(*
SPDX-FileCopyrightText: © 2026 Oleksandr Tiutyk <trofimich@gmail.com>
SPDX-License-Identifier: MIT
License: https://opensource.org/license/mit
*)

(*!
<summary>Serializes live PLC structures to JSON and restores them from JSON.</summary>
<description>
Supports live PLC structures with native type information; dynamically created structures are not supported.
ByVarInfo methods require an explicit PVOID address; descriptor ByteAddress is ignored to preserve pointer width.
Application method calls and property access belong to one owner task per instance. Instances are not
thread-safe and do not support reentry: a callback must not call methods or access properties of the
serializer whose operation is still active, directly or indirectly. Use a separate instance and separate
buffers for another task or nested conversion. Ownership is a caller precondition, not a runtime check or
lock; Try does not make an ownership violation safe or guarantee its detection as FALSE. Keep source data
stable and destination storage exclusive for the entire call, including callbacks. Separate serializer
instances do not synchronize shared application data. Stateful extenders require their own ownership
discipline; sharing an extender must not introduce concurrent state access. Borrows input, output and optional
callbacks for each call. Throwing methods report invalid arguments and native failures through framework
exceptions. Try methods return FALSE directly for rejected arguments or reported native failures and contain
exceptions from native calls or callbacks; partial effects are not rolled back. Try methods use the shared
native conversion helpers, not overrides of the throwing methods or their protected helpers. JSON text uses
native UTF-8 encoding; capacity and copy sizes count bytes. Instances must not be copied by value. The caller
provides cyclic-task exception cleanup and RaiseIfAllocationFailed at the task boundary, outside Try and
recoverable handlers. Try methods do not clear terminal allocation state. Ownership examples and future
shared-service guidance: Guides/JsonAndEventLoggerOwnership.md in the repository.
</description>
*)

{attribute 'no_explicit_call' := 'Direct call is not allowed'}
FUNCTION_BLOCK AutomaticJsonSerializer EXTENDS TOF_Core.Object
VAR_STAT
	//! <summary>Class name shared by all instances of this function block.</summary>
	{attribute 'hide'} 
	_ClassName : STRING := __POUNAME();
END_VAR
VAR
	_JsonSaxWriter : Tc3_JsonXml.FB_JsonSaxWriter;
	_JsonDataTypeWriter : Tc3_JsonXml.FB_JsonReadWriteDatatype;
END_VAR

(*!
<summary>Provides the concrete serializer class name.</summary>
<description>Borrows read-only instance storage that remains valid for the instance lifetime.</description>
*)
{attribute 'monitoring' := 'call'}
PROPERTY ClassName : REFERENCE TO STRING
GET
ClassName REF= _ClassName;
END_GET
END_PROPERTY

(*!
<summary>Serializes a PLC structure into caller-owned JSON storage.</summary>
<description>
Uses native symbol lookup for the source type; dynamically created structures are not supported. Single-field
structures have native lookup limitations; use ByVarInfo to supply the type explicitly. Borrows
source, destination and optional extender for the call. The destination must be writable and have at least
JSON_DOCUMENT capacity. Invalid source arguments and reported native failures raise framework exceptions;
extender exceptions propagate. Output and callback effects are not rolled back on failure. Exception transport
and cleanup require the caller's cyclic-task boundary. CopyDocument returning zero or a nonzero HRESULT raises
an exception; jsonSize is not usable on failure.
</description>
<param name="sourceStructure">Live PLC structure with type information available to native symbol lookup.</param>
<param name="extender">
Optional callback invoked before and after writing the structure value; zero skips both calls.
</param>
<param name="targetJson">Writable output storage with at least 25000 bytes of text capacity plus the terminator.</param>
<param name="jsonSize">
Byte count reported by CopyDocument, including the terminator on a successful copy; use only after normal
completion.
</param>
*)
METHOD Serialize
VAR_INPUT
	sourceStructure : ANY;
	extender : IJsonExtender := 0;
END_VAR
VAR_IN_OUT
	targetJson : TOF_Core.JSON_DOCUMENT;
END_VAR
VAR_OUTPUT
	jsonSize : UDINT; 
END_VAR
InternalSerialize(
	sourceStructure := sourceStructure,
	extender := extender,
	targetJson := targetJson,
	jsonSize => jsonSize
);
END_METHOD

(*!
<summary>Serializes a PLC structure described by VAR_INFO into caller-owned JSON storage.</summary>
<description>
The descriptor type and byte-aligned size must match sourceStructureAddress. ByteAddress is ignored.
Dynamically created structures are not supported. Borrows source, destination and optional extender for the call. The
destination must be writable and have at least JSON_DOCUMENT capacity. Invalid source arguments and reported
native failures raise framework exceptions; extender exceptions propagate. Output and callback effects are not
rolled back on failure. Exception transport and cleanup require the caller's cyclic-task boundary.
CopyDocument returning zero or a nonzero HRESULT raises an exception; jsonSize is not usable on failure.
</description>
<param name="sourceStructureAddress">
Required address from ADR of the live source structure, borrowed for this call. Must match the descriptor.
Zero is rejected; no address is recovered from ByteAddress or ByteOffset.
</param>
<param name="sourceStructureVarInfo">
Descriptor whose TypeName and BitSize describe the source structure; ByteAddress is ignored.
</param>
<param name="extender">
Optional callback invoked before and after writing the structure value; zero skips both calls.
</param>
<param name="targetJson">Writable output storage with at least 25000 bytes of text capacity plus the terminator.</param>
<param name="jsonSize">
Byte count reported by CopyDocument, including the terminator on a successful copy; use only after normal
completion.
</param>
*)
METHOD SerializeByVarInfo
VAR_INPUT
	sourceStructureVarInfo : __SYSTEM.VAR_INFO;
	sourceStructureAddress : PVOID;
	extender : IJsonExtender := 0;
END_VAR
VAR_IN_OUT
	targetJson : TOF_Core.JSON_DOCUMENT;
END_VAR
VAR_OUTPUT
	jsonSize : UDINT; 
END_VAR
VAR
	formattedExceptionMessage : TOF_Core.ERROR_MESSAGE;

	
	errorCode : HRESULT;
END_VAR
IF sourceStructureAddress = TOF_Core.Memory.NULL_ADDRESS THEN
	TOF_Core.Exceptions.ThrowArgumentNotSpecified(
		sourceNamespaceName := NamespaceName,
		sourceClassName := ClassName,
		sourcePOUName := __POUNAME(),
		sourcePosition := __POSITION(),
		argumentName := 'sourceStructureAddress'
	);
END_IF

IF sourceStructureVarInfo.TypeClass <> __SYSTEM.TYPE_CLASS.TYPE_USERDEF THEN
	TOF_Core.Exceptions.ThrowArgumentTypeClassNotSupported(
		sourceNamespaceName := NamespaceName,
		sourceClassName := ClassName,
		sourcePOUName := __POUNAME(),
		sourcePosition := __POSITION(),
		argumentName := 'sourceStructureVarInfo',
		argumentType := sourceStructureVarInfo.TypeClass
	);
END_IF

// VAR_INFO sizes are in bits; the caller supplies a byte-aligned structure descriptor.
IF NOT writeStructureJson(
	structureTypeName := sourceStructureVarInfo.TypeName,
	structureAddress := sourceStructureAddress,
	structureSize := TO_UDINT(sourceStructureVarInfo.BitSize / 8),
	extender := extender,
	targetJson := targetJson,
	jsonSize => jsonSize,
	errorCode => errorCode,
	errorMessage => formattedExceptionMessage
)
THEN
	TOF_Core.Exceptions.ThrowStandard(
		sourceNamespaceName := NamespaceName,
		sourceClassName := ClassName,
		sourcePOUName := __POUNAME(),
		sourcePosition := __POSITION(),
		message := formattedExceptionMessage,
		errorCode := TO_UDINT(errorCode)
	);
END_IF
END_METHOD

{attribute 'monitoring' := 'call'}
(*!
<summary>Gets or sets the native writer's maximum number of fractional decimal places.</summary>
<description>
The native writer determines which DINT values it supports; this property does not clamp the value. The setter
requires a zero HRESULT from SetMaxDecimalPlaces. A nonzero HRESULT raises a framework exception because
assignment has no failure result. The native error code is retained in the exception. No rollback of the
native setting is guaranteed on failure; the getter reads the writer's current setting. The caller handles the
exception and provides cyclic-task exception cleanup and the terminal allocation-failure boundary.
</description>
*)
PROPERTY DecimalPlaces : DINT
GET
DecimalPlaces := _JsonSaxWriter.GetMaxDecimalPlaces();
END_GET
SET
VAR
	errorCode : HRESULT;
END_VAR
errorCode := _JsonSaxWriter.SetMaxDecimalPlaces(decimalPlaces := DecimalPlaces);

IF errorCode <> TOF_Core.SignedInt32.ZERO THEN
	TOF_Core.Exceptions.ThrowStandard(
		sourceNamespaceName := NamespaceName,
		sourceClassName := ClassName,
		sourcePOUName := __POUNAME(),
		sourcePosition := __POSITION(),
		message := "Can't set JSON writer decimal places",
		errorCode := TO_UDINT(errorCode)
	);
END_IF
END_SET
END_PROPERTY

(*!
<summary>Populates a PLC structure from JSON using the type supplied by VAR_INFO.</summary>
<description>
TypeName and byte-aligned BitSize must describe the live, writable structure at targetStructureAddress.
ByteAddress is ignored. Uses the supplied TypeName directly, avoiding ambiguous address-based type lookup
for single-field structures. The type
must be available to the native JSON converter; support for dynamically created structures is not implied.
Borrows the JSON and destination for this call. A zero address, an unsupported type class or a reported native
conversion failure raises a framework exception. Conversion requires both a TRUE SetSymbolFromJson result and
a zero HRESULT. Destination fields may already have changed on failure; writes are not rolled back. The caller
provides cyclic-task exception cleanup and the terminal allocation-failure boundary.
</description>
<param name="json">JSON text to read without modification.</param>
<param name="targetStructureAddress">
Required address from ADR of the live target structure, borrowed for this call. Must match the descriptor.
Zero is rejected; no address is recovered from ByteAddress or ByteOffset.
</param>
<param name="targetStructureVarInfo">
Consistent descriptor of the destination structure, including its explicit TypeName.
</param>
*)
METHOD DeserializeByVarInfo
VAR_IN_OUT CONSTANT
	json : TOF_Core.JSON_DOCUMENT;	
END_VAR
VAR_INPUT
	targetStructureVarInfo : __SYSTEM.VAR_INFO;
	targetStructureAddress : PVOID;
END_VAR
VAR
	
	errorCode : HRESULT;
END_VAR
IF targetStructureAddress = TOF_Core.Memory.NULL_ADDRESS THEN
	TOF_Core.Exceptions.ThrowArgumentNotSpecified(
		sourceNamespaceName := NamespaceName,
		sourceClassName := ClassName,
		sourcePOUName := __POUNAME(),
		sourcePosition := __POSITION(),
		argumentName := 'targetStructureAddress'
	);
END_IF

IF targetStructureVarInfo.TypeClass <> __SYSTEM.TYPE_CLASS.TYPE_USERDEF THEN
	TOF_Core.Exceptions.ThrowArgumentTypeClassNotSupported(
		sourceNamespaceName := NamespaceName,
		sourceClassName := ClassName,
		sourcePOUName := __POUNAME(),
		sourcePosition := __POSITION(),
		argumentName := 'targetStructureVarInfo',
		argumentType := targetStructureVarInfo.TypeClass
	);
END_IF

// VAR_INFO sizes are in bits; the caller supplies a byte-aligned structure descriptor.
IF NOT readStructureJson(
	json := json,
	structureTypeName := targetStructureVarInfo.TypeName,
	structureAddress := targetStructureAddress,
	structureSize := TO_UDINT(targetStructureVarInfo.BitSize / 8),
	errorCode => errorCode
)
THEN
	TOF_Core.Exceptions.ThrowStandard(
		sourceNamespaceName := NamespaceName,
		sourceClassName := ClassName,
		sourcePOUName := __POUNAME(),
		sourcePosition := __POSITION(),
		message := "Can't fill target structure by specified json document",
		errorCode := TO_UDINT(errorCode)
	);
END_IF
END_METHOD

(*!
<summary>Populates a PLC structure from JSON using native address-based type lookup.</summary>
<description>
Borrows the JSON and a live, writable structure for the call; dynamically created structures are not
supported. Native type lookup has limitations for single-field structures. Invalid arguments, reported lookup
failures, a FALSE SetSymbolFromJson result or a nonzero conversion HRESULT raise framework exceptions.
Destination fields may already have changed on failure; writes are not rolled back. The caller provides
cyclic-task exception cleanup and the terminal allocation-failure boundary.
</description>
<param name="json">JSON text to read without modification.</param>
<param name="targetStructure">
Live destination structure with type information available to native symbol lookup.
</param>
*)
METHOD Deserialize
VAR_IN_OUT CONSTANT
	json : TOF_Core.JSON_DOCUMENT;	
END_VAR
VAR_INPUT
	targetStructure : ANY;
END_VAR
InternalDeserialize(json := json, targetStructure := targetStructure);
END_METHOD

(*!
<summary>Serializes a structure using its ANY descriptor and native symbol lookup.</summary>
<description>
The descriptor must identify a live structure with matching address and size; dynamically created structures
are not supported. Native address lookup has limitations for single-field structures. Borrows source,
destination and optional extender for the call. The destination must be writable and have at least
JSON_DOCUMENT capacity. Invalid source arguments and reported native failures raise framework exceptions;
extender exceptions propagate. Output and callback effects are not rolled back on failure. Overrides must
preserve destination capacity and borrowing requirements. This protected hook serves the throwing ANY API;
TrySerialize does not dispatch through it. Exception transport and cleanup require the caller's
cyclic-task boundary. CopyDocument returning zero or a nonzero HRESULT raises an exception; jsonSize is not
usable on failure.
</description>
<param name="sourceStructure">ANY descriptor for the source structure.</param>
<param name="extender">
Optional callback invoked before and after writing the structure value; zero skips both calls.
</param>
<param name="targetJson">Writable output storage with at least 25000 bytes of text capacity plus the terminator.</param>
<param name="jsonSize">
Byte count reported by CopyDocument, including the terminator on a successful copy; use only after normal
completion.
</param>
*)
METHOD PROTECTED InternalSerialize
VAR_INPUT
	sourceStructure : __SYSTEM.AnyType;
	extender : IJsonExtender := 0;
END_VAR
VAR_IN_OUT
	targetJson : TOF_Core.JSON_DOCUMENT;
END_VAR
VAR_OUTPUT
	jsonSize : UDINT; 
END_VAR
VAR
	formattedExceptionMessage : TOF_Core.ERROR_MESSAGE;

	
	structureTypeName : STRING;	 
	errorCode : HRESULT;
END_VAR
IF sourceStructure.pValue = TOF_Core.Memory.NULL_ADDRESS THEN
	TOF_Core.Exceptions.ThrowArgumentNotSpecified(
		sourceNamespaceName := NamespaceName,
		sourceClassName := ClassName,
		sourcePOUName := __POUNAME(),
		sourcePosition := __POSITION(),
		argumentName := 'sourceStructure'
	);
END_IF

IF sourceStructure.TypeClass <> __SYSTEM.TYPE_CLASS.TYPE_USERDEF THEN
	TOF_Core.Exceptions.ThrowArgumentTypeClassNotSupported(
		sourceNamespaceName := NamespaceName,
		sourceClassName := ClassName,
		sourcePOUName := __POUNAME(),
		sourcePosition := __POSITION(),
		argumentName := 'sourceStructure',
		argumentType := sourceStructure.TypeClass
	);
END_IF

structureTypeName := _JsonDataTypeWriter.GetDatatypeNameByAddress(
	nData := TO_UDINT(sourceStructure.diSize),
	pData := sourceStructure.pValue,
	hrErrorCode => errorCode
);

IF errorCode <> TOF_Core.SignedInt32.ZERO THEN
	TOF_Core.Exceptions.ThrowStandard(
		sourceNamespaceName := NamespaceName,
		sourceClassName := ClassName,
		sourcePOUName := __POUNAME(),
		sourcePosition := __POSITION(),
		message := "Can't get structure type of the source structure",
		errorCode := TO_UDINT(errorCode)
	);
END_IF

IF NOT writeStructureJson(
	structureTypeName := structureTypeName,
	structureAddress := sourceStructure.pValue,
	structureSize := TO_UDINT(sourceStructure.diSize),
	extender := extender,
	targetJson := targetJson,
	jsonSize => jsonSize,
	errorCode => errorCode,
	errorMessage => formattedExceptionMessage
)
THEN
	TOF_Core.Exceptions.ThrowStandard(
		sourceNamespaceName := NamespaceName,
		sourceClassName := ClassName,
		sourcePOUName := __POUNAME(),
		sourcePosition := __POSITION(),
		message := formattedExceptionMessage,
		errorCode := TO_UDINT(errorCode)
	);
END_IF
END_METHOD

(*!
<summary>Deserializes JSON into the structure identified by an ANY descriptor.</summary>
<description>
The descriptor must identify a live, writable structure with matching address and size; dynamically created
structures are not supported. Native address-based type lookup has limitations for single-field structures.
Borrows the JSON and destination for the call. Invalid arguments, reported lookup failures, a FALSE
SetSymbolFromJson result or a nonzero conversion HRESULT raise framework exceptions. Partial destination
writes are not rolled back. Overrides must preserve borrowing and failure reporting requirements. This
protected hook serves the throwing ANY API; TryDeserialize does not dispatch through it. The caller
provides cyclic-task exception cleanup and the terminal allocation-failure boundary.
</description>
<param name="json">JSON text to read without modification.</param>
<param name="targetStructure">ANY descriptor for the live destination structure.</param>
*)
METHOD PROTECTED InternalDeserialize
VAR_IN_OUT CONSTANT
	json : TOF_Core.JSON_DOCUMENT;	
END_VAR
VAR_INPUT
	targetStructure : __SYSTEM.AnyType;
END_VAR
VAR
	
	structureTypeName : STRING;	 
	errorCode : HRESULT;
END_VAR
IF targetStructure.pValue = TOF_Core.Memory.NULL_ADDRESS THEN
	TOF_Core.Exceptions.ThrowArgumentNotSpecified(
		sourceNamespaceName := NamespaceName,
		sourceClassName := ClassName,
		sourcePOUName := __POUNAME(),
		sourcePosition := __POSITION(),
		argumentName := 'targetStructure'
	);
END_IF

IF targetStructure.TypeClass <> __SYSTEM.TYPE_CLASS.TYPE_USERDEF THEN
	TOF_Core.Exceptions.ThrowArgumentTypeClassNotSupported(
		sourceNamespaceName := NamespaceName,
		sourceClassName := ClassName,
		sourcePOUName := __POUNAME(),
		sourcePosition := __POSITION(),
		argumentName := 'targetStructure',
		argumentType := targetStructure.TypeClass
	);
END_IF

structureTypeName := _JsonDataTypeWriter.GetDatatypeNameByAddress(
	nData := TO_UDINT(targetStructure.diSize),
	pData := targetStructure.pValue,
	hrErrorCode => errorCode
);

IF errorCode <> TOF_Core.SignedInt32.ZERO THEN
	TOF_Core.Exceptions.ThrowStandard(
		sourceNamespaceName := NamespaceName,
		sourceClassName := ClassName,
		sourcePOUName := __POUNAME(),
		sourcePosition := __POSITION(),
		message := "Can't get structure type of the target structure",
		errorCode := TO_UDINT(errorCode)
	);
END_IF

IF NOT readStructureJson(
	json := json,
	structureTypeName := structureTypeName,
	structureAddress := targetStructure.pValue,
	structureSize := TO_UDINT(targetStructure.diSize),
	errorCode => errorCode
)
THEN
	TOF_Core.Exceptions.ThrowStandard(
		sourceNamespaceName := NamespaceName,
		sourceClassName := ClassName,
		sourcePOUName := __POUNAME(),
		sourcePosition := __POSITION(),
		message := "Can't fill target structure by specified json document",
		errorCode := TO_UDINT(errorCode)
	);
END_IF
END_METHOD

(*!
<summary>Provides the compiler-initialized library namespace.</summary>
<description>Borrows read-only library storage; no allocation or ownership transfer occurs.</description>
*)
{attribute 'monitoring' := 'call'}
PROPERTY NamespaceName : REFERENCE TO STRING
GET
NamespaceName REF= CurrentNamespace.Name;
END_GET
END_PROPERTY

(*!
<summary>Reads JSON into a validated structure and reports the native conversion result.</summary>
<description>
Callers validate the descriptor before entry. Borrows the JSON, type name and destination for this call.
Returns FALSE for a native FALSE result or nonzero HRESULT without creating exceptions. Native exceptions
propagate to the throwing caller or the public Try boundary. Checks fatal allocation state before conversion
and before reporting success, raising a contained terminal failure without constructing an exception object.
The Try boundary converts that failure to FALSE. Partial destination writes are not rolled back.
</description>
<param name="json">JSON text to read without modification.</param>
<param name="structureTypeName">Native type name matching the destination structure.</param>
<param name="structureAddress">Address of the validated writable destination.</param>
<param name="structureSize">Destination structure size in bytes.</param>
<param name="errorCode">Native conversion HRESULT, interpreted together with the BOOL result.</param>
*)
METHOD PRIVATE readStructureJson : BOOL
VAR_IN_OUT CONSTANT
	json : TOF_Core.JSON_DOCUMENT;
	structureTypeName : STRING;
END_VAR
VAR_INPUT
	structureAddress : PVOID;
	structureSize : UDINT;
END_VAR
VAR_OUTPUT
	errorCode : HRESULT;
END_VAR
TOF_Core.DynamicMemoryManager.RaiseIfAllocationFailed();

IF NOT _JsonDataTypeWriter.SetSymbolFromJson(
		sJson := json,
		sDatatype := structureTypeName,
		nData := structureSize,
		pData := structureAddress,
		hrErrorCode => errorCode
	)
	OR_ELSE errorCode <> TOF_Core.SignedInt32.ZERO
THEN
	RETURN;
END_IF

TOF_Core.DynamicMemoryManager.RaiseIfAllocationFailed();
readStructureJson := TRUE;
END_METHOD

(*!
<summary>Reports the complete instance size in bytes.</summary>
<description>Uses XSIZEOF; separately allocated native resources are not included.</description>
*)
{attribute 'monitoring' := 'call'}
PROPERTY SelfSize : ULINT
GET
SelfSize := XSIZEOF(THIS^);
END_GET
END_PROPERTY

{attribute 'TcRpcEnable':='1'}
(*!
<summary>Attempts to serialize a PLC structure to JSON.</summary>
<description>
Returns FALSE directly for a null address, an unsupported type class or a reported native failure, including a
zero CopyDocument result, without creating a framework exception. Contains native and callback exceptions.
Uses the shared conversion helper rather than the protected throwing hook. Use JSON and jsonSize only on TRUE;
partial writes and callback effects are not rolled back. Each subsequent conversion attempts to reset the
writer before callbacks. Borrows live source and writable destination storage. Does not clear terminal allocation state; the
caller provides exception cleanup and RaiseIfAllocationFailed at the task boundary outside Try and recoverable
handlers. Returns FALSE when fatal allocation state is observed on entry or after nested calls; a contained
allocation failure is not a successful conversion. The application-wide latch remains set.
</description>
<param name="sourceStructure">
Live PLC structure supported by native symbol lookup; dynamically created structures are not supported.
Single-field structures have native lookup limitations; use ByVarInfo to supply the type explicitly.
</param>
<param name="extender">
Optional callback invoked before and after writing the structure value; borrowed for the call.
</param>
<param name="targetJson">
Writable output storage with at least 25000 bytes of text capacity plus the terminator; borrowed for the call.
</param>
<param name="jsonSize">
Byte count reported by CopyDocument, including the terminator on a successful copy; use only on TRUE.
</param>
*)
METHOD TrySerialize : BOOL
VAR_INPUT
	sourceStructure : ANY;
	extender : IJsonExtender := 0;
END_VAR
VAR_IN_OUT
	targetJson : TOF_Core.JSON_DOCUMENT;
END_VAR
VAR_OUTPUT
	jsonSize : UDINT; 
END_VAR
VAR
	structureTypeName : STRING;
	errorCode : HRESULT;
END_VAR
__TRY

	IF TOF_Core.DynamicMemoryManager.HasAllocationFailed THEN
		RETURN;
	END_IF

	IF sourceStructure.pValue = TOF_Core.Memory.NULL_ADDRESS
		OR_ELSE sourceStructure.TypeClass <> __SYSTEM.TYPE_CLASS.TYPE_USERDEF
	THEN
		RETURN;
	END_IF

	structureTypeName := _JsonDataTypeWriter.GetDatatypeNameByAddress(
		nData := TO_UDINT(sourceStructure.diSize),
		pData := sourceStructure.pValue,
		hrErrorCode => errorCode
	);

	IF errorCode <> TOF_Core.SignedInt32.ZERO THEN
		RETURN;
	END_IF

	TrySerialize := writeStructureJson(
		structureTypeName := structureTypeName,
		structureAddress := sourceStructure.pValue,
		structureSize := TO_UDINT(sourceStructure.diSize),
		extender := extender,
		targetJson := targetJson,
		jsonSize => jsonSize
	);

	IF TOF_Core.DynamicMemoryManager.HasAllocationFailed THEN
		TrySerialize := FALSE;
	END_IF

__CATCH
	TrySerialize := FALSE;
__ENDTRY
END_METHOD

(*!
<summary>Attempts to serialize a PLC structure to JSON.</summary>
<description>
Returns FALSE directly for a null address, an unsupported type class or a reported native failure, including a
zero CopyDocument result, without creating a framework exception. Contains native and callback exceptions.
Uses the shared conversion helper rather than the throwing ByVarInfo method. Use JSON and jsonSize only on
TRUE; partial writes and callback effects are not rolled back. Each subsequent conversion attempts to reset
the writer before callbacks. Borrows live source and writable destination storage. Does not clear terminal allocation
state; the caller provides exception cleanup and RaiseIfAllocationFailed at the task boundary outside Try and
recoverable handlers. Returns FALSE when fatal allocation state is observed on entry or after nested calls; a contained
allocation failure is not a successful conversion. The application-wide latch remains set.
</description>
<param name="sourceStructureAddress">
Required address from ADR of the live source structure, borrowed for this call. Must match the descriptor.
Zero is rejected; no address is recovered from ByteAddress or ByteOffset.
</param>
<param name="sourceStructureVarInfo">
Descriptor with matching TypeName and byte-aligned BitSize for sourceStructureAddress; ByteAddress is ignored.
Dynamically created structures are not supported.
</param>
<param name="extender">
Optional callback invoked before and after writing the structure value; borrowed for the call.
</param>
<param name="targetJson">
Writable output storage with at least 25000 bytes of text capacity plus the terminator; borrowed for the call.
</param>
<param name="jsonSize">
Byte count reported by CopyDocument, including the terminator on a successful copy; use only on TRUE.
</param>
*)
METHOD TrySerializeByVarInfo : BOOL
VAR_INPUT
	sourceStructureVarInfo : __SYSTEM.VAR_INFO;
	sourceStructureAddress : PVOID;
	extender : IJsonExtender := 0;
END_VAR
VAR_IN_OUT
	targetJson : TOF_Core.JSON_DOCUMENT;
END_VAR
VAR_OUTPUT
	jsonSize : UDINT; 
END_VAR
__TRY

	IF TOF_Core.DynamicMemoryManager.HasAllocationFailed THEN
		RETURN;
	END_IF

	IF sourceStructureAddress = TOF_Core.Memory.NULL_ADDRESS
		OR_ELSE sourceStructureVarInfo.TypeClass <> __SYSTEM.TYPE_CLASS.TYPE_USERDEF
	THEN
		RETURN;
	END_IF

	// VAR_INFO sizes are in bits; the descriptor must be byte-aligned.
	TrySerializeByVarInfo := writeStructureJson(
		structureTypeName := sourceStructureVarInfo.TypeName,
		structureAddress := sourceStructureAddress,
		structureSize := TO_UDINT(sourceStructureVarInfo.BitSize / 8),
		extender := extender,
		targetJson := targetJson,
		jsonSize => jsonSize
	);

	IF TOF_Core.DynamicMemoryManager.HasAllocationFailed THEN
		TrySerializeByVarInfo := FALSE;
	END_IF

__CATCH
	TrySerializeByVarInfo := FALSE;
__ENDTRY
END_METHOD

(*!
<summary>Attempts to populate a PLC structure from JSON using the type supplied by VAR_INFO.</summary>
<description>
Uses the supplied TypeName directly without address-based type lookup. TypeName and byte-aligned BitSize must
describe the live, writable structure at targetStructureAddress, with its type available to the native converter.
ByteAddress is ignored.
Returns FALSE directly for a null address, an unsupported type class, a FALSE native conversion result or a
nonzero HRESULT, without creating a framework exception. Contains native exceptions. Uses the shared
conversion helper rather than the throwing ByVarInfo method. Partial destination writes are not rolled back.
Borrows the JSON and destination for this call. Does not clear terminal allocation state; the caller provides
exception cleanup and RaiseIfAllocationFailed at the task boundary outside Try and recoverable handlers.
Returns FALSE when fatal allocation state is observed on entry or after nested calls; a contained
allocation failure is not a successful conversion. The application-wide latch remains set.
</description>
<param name="json">JSON text to read without modification.</param>
<param name="targetStructureAddress">
Required address from ADR of the live target structure, borrowed for this call. Must match the descriptor.
Zero is rejected; no address is recovered from ByteAddress or ByteOffset.
</param>
<param name="targetStructureVarInfo">
Consistent descriptor of the destination structure, including its explicit TypeName.
</param>
*)
METHOD TryDeserializeByVarInfo : BOOL
VAR_IN_OUT CONSTANT
	json : TOF_Core.JSON_DOCUMENT;	
END_VAR
VAR_INPUT
	targetStructureVarInfo : __SYSTEM.VAR_INFO;
	targetStructureAddress : PVOID;
END_VAR
__TRY

	IF TOF_Core.DynamicMemoryManager.HasAllocationFailed THEN
		RETURN;
	END_IF

	IF targetStructureAddress = TOF_Core.Memory.NULL_ADDRESS
		OR_ELSE targetStructureVarInfo.TypeClass <> __SYSTEM.TYPE_CLASS.TYPE_USERDEF
	THEN
		RETURN;
	END_IF

	// VAR_INFO sizes are in bits; the descriptor must be byte-aligned.
	TryDeserializeByVarInfo := readStructureJson(
		json := json,
		structureTypeName := targetStructureVarInfo.TypeName,
		structureAddress := targetStructureAddress,
		structureSize := TO_UDINT(targetStructureVarInfo.BitSize / 8)
	);

	IF TOF_Core.DynamicMemoryManager.HasAllocationFailed THEN
		TryDeserializeByVarInfo := FALSE;
	END_IF

__CATCH
	TryDeserializeByVarInfo := FALSE;
__ENDTRY
END_METHOD

(*!
<summary>Attempts to populate a PLC structure from JSON.</summary>
<description>
Uses native address-based type lookup, with its limitations for single-field structures; dynamically created
structures are not supported. Returns FALSE directly for a null address, an unsupported type class, a reported
lookup failure, a FALSE native conversion result or a nonzero conversion HRESULT, without creating a framework
exception. Contains native exceptions. Uses the shared conversion helper rather than the protected throwing
hook. Partial destination writes are not rolled back. Borrows JSON and live, writable destination storage for
this call. Does not clear terminal allocation state; the caller provides exception cleanup and
RaiseIfAllocationFailed at the task boundary outside Try and recoverable handlers.
Returns FALSE when fatal allocation state is observed on entry or after nested calls; a contained
allocation failure is not a successful conversion. The application-wide latch remains set.
</description>
<param name="json">JSON text to read without modification.</param>
<param name="targetStructure">
Live destination structure with type information available to native symbol lookup.
</param>
*)
METHOD TryDeserialize : BOOL
VAR_IN_OUT CONSTANT
	json : TOF_Core.JSON_DOCUMENT;	
END_VAR
VAR_INPUT
	targetStructure : ANY;
END_VAR
VAR
	structureTypeName : STRING;
	errorCode : HRESULT;
END_VAR
__TRY

	IF TOF_Core.DynamicMemoryManager.HasAllocationFailed THEN
		RETURN;
	END_IF

	IF targetStructure.pValue = TOF_Core.Memory.NULL_ADDRESS
		OR_ELSE targetStructure.TypeClass <> __SYSTEM.TYPE_CLASS.TYPE_USERDEF
	THEN
		RETURN;
	END_IF

	structureTypeName := _JsonDataTypeWriter.GetDatatypeNameByAddress(
		nData := TO_UDINT(targetStructure.diSize),
		pData := targetStructure.pValue,
		hrErrorCode => errorCode
	);

	IF errorCode <> TOF_Core.SignedInt32.ZERO THEN
		RETURN;
	END_IF

	TryDeserialize := readStructureJson(
		json := json,
		structureTypeName := structureTypeName,
		structureAddress := targetStructure.pValue,
		structureSize := TO_UDINT(targetStructure.diSize)
	);

	IF TOF_Core.DynamicMemoryManager.HasAllocationFailed THEN
		TryDeserialize := FALSE;
	END_IF

__CATCH
	TryDeserialize := FALSE;
__ENDTRY
END_METHOD

(*!
<summary>Writes a validated structure and optional extensions to caller-owned JSON storage.</summary>
<description>
Callers validate the structure descriptor before entry. Borrows all arguments for this call and resets the
writer before invoking callbacks. A nonzero ResetDocument HRESULT returns FALSE before any hook or copy.
Returns FALSE for reported native failures without creating exceptions; native or callback exceptions propagate
to the throwing caller or the public Try boundary. Checks fatal allocation state before native work, after
successful native steps and after each hook. A contained terminal failure is raised again without allocating
an exception object; the Try boundary converts it to FALSE. No output, writer or callback effects are rolled
back. Each later write attempts to reset the writer again. On FALSE, errorMessage describes the failed native
step and errorCode retains its HRESULT without substitution.
</description>
<param name="structureTypeName">Native type name matching the live source structure.</param>
<param name="structureAddress">Address of the validated source structure.</param>
<param name="structureSize">Source structure size in bytes.</param>
<param name="extender">Optional callbacks around the structure value.</param>
<param name="targetJson">Writable storage with JSON_DOCUMENT capacity, including its terminator.</param>
<param name="jsonSize">Copied byte count including the terminator; meaningful only on TRUE.</param>
<param name="errorCode">Native HRESULT of the failed step on FALSE.</param>
<param name="errorMessage">Diagnostic for the failed step on FALSE.</param>
*)
METHOD PRIVATE writeStructureJson : BOOL
VAR_IN_OUT CONSTANT
	structureTypeName : STRING;
END_VAR
VAR_INPUT
	structureAddress : PVOID;
	structureSize : UDINT;
	extender : IJsonExtender;
END_VAR
VAR_IN_OUT
	targetJson : TOF_Core.JSON_DOCUMENT;
END_VAR
VAR_OUTPUT
	jsonSize : UDINT;
	errorCode : HRESULT;
	errorMessage : WSTRING(255);
END_VAR
TOF_Core.DynamicMemoryManager.RaiseIfAllocationFailed();
errorCode := _JsonSaxWriter.ResetDocument();
TOF_Core.DynamicMemoryManager.RaiseIfAllocationFailed();

IF errorCode <> TOF_Core.SignedInt32.ZERO THEN
	errorMessage := "Can't reset JSON writer before structure serialization";
	RETURN;
END_IF

IF extender <> 0 THEN
	extender.WritePrefix(jsonSaxWriter := _JsonSaxWriter);
	TOF_Core.DynamicMemoryManager.RaiseIfAllocationFailed();
END_IF

IF NOT _JsonDataTypeWriter.AddJsonValueFromSymbol(
		fbWriter := _JsonSaxWriter,
		sDatatype := structureTypeName,
		nData := structureSize,
		pData := structureAddress,
		hrErrorCode => errorCode
	)
	OR_ELSE errorCode <> TOF_Core.SignedInt32.ZERO
THEN
	errorMessage := TOF_Core.WideStrings.Concat255(
		"Can't generate JSON representation from the symbol of type '",
		TO_WSTRING(structureTypeName),
		"'"
	);
	RETURN;
END_IF

TOF_Core.DynamicMemoryManager.RaiseIfAllocationFailed();

IF extender <> 0 THEN
	extender.WriteSuffix(jsonSaxWriter := _JsonSaxWriter);
	TOF_Core.DynamicMemoryManager.RaiseIfAllocationFailed();
END_IF

jsonSize := _JsonSaxWriter.CopyDocument(
	pDoc := targetJson,
	nDoc := SIZEOF(targetJson),
	hrErrorCode => errorCode
);

IF jsonSize = TOF_Core.UnsignedInt32.MIN_VALUE OR_ELSE errorCode <> TOF_Core.SignedInt32.ZERO THEN
	errorMessage := TOF_Core.WideStrings.Concat255(
		"Can't fill JSON from the symbol of type '",
		TO_WSTRING(structureTypeName),
		"'"
	);
	RETURN;
END_IF

TOF_Core.DynamicMemoryManager.RaiseIfAllocationFailed();
writeStructureJson := TRUE;
END_METHOD

END_FUNCTION_BLOCK

(* stored: Version 1.1.0.1
   POU AutomaticJsonSerializer: Id {a4623321-e5e2-4514-b5b7-6f50c93efdb9}, SpecialFunc None
   Folder Service memebers: Id {ac3ba484-d0b1-4d7e-b557-cd243c8b8997}
   Property ClassName: Id {0ef034e0-c59c-400d-8910-5199a1e43c28}
   Get Get: Id {7d8e441f-d9e1-4fe6-a84f-2d3a88ae1b83}
   Method Serialize: Id {defd30bb-3636-4b3d-a29d-4ee5f3966212}
   Method SerializeByVarInfo: Id {d6f652b9-17a4-4ec4-936c-676a73e01a2d}
   Property DecimalPlaces: Id {856a998f-c63b-4bfb-be2d-ebc0ce7cf745}
   Get Get: Id {94eff383-c1b9-45b7-8cbb-da0c6c3a2aac}
   Set Set: Id {e5e3c1bb-4425-43f2-a416-2b4fee3a3ddc}
   Method DeserializeByVarInfo: Id {3b0559f7-3cc9-4407-b03c-9992acf72583}
   Method Deserialize: Id {b53042c3-1eea-4151-a973-f56939241dea}
   Method InternalSerialize: Id {828ddc06-4e4b-4f22-bd8f-3234f73fd728}
   Method InternalDeserialize: Id {cd668581-fbff-4bb3-b0d3-914c47132fdf}
   Property NamespaceName: Id {7371ecef-1936-4268-af0d-813ed5877183}
   Get Get: Id {a712aceb-e580-4469-b321-74f0e6ab0c97}
   Method readStructureJson: Id {e9710e74-d168-4bec-aecb-ed84a0f769b4}
   Property SelfSize: Id {4e2cc4a2-86a6-48cc-a757-58f1b82e3903}
   Get Get: Id {3c9a353a-dae3-4a6a-8486-44c6e5bd0b57}
   Method TrySerialize: Id {35373f3b-1087-4a79-950c-0b141211bf99}
   Method TrySerializeByVarInfo: Id {486e285a-fcfe-44f3-9023-743f121d8975}
   Method TryDeserializeByVarInfo: Id {25972cd3-eceb-4afa-aeb2-ef7585c39b37}
   Method TryDeserialize: Id {b5b62249-7ff4-4c95-ba2a-e43e9757d053}
   Method writeStructureJson: Id {b6245462-dfce-45a0-a956-f50e59e6d73a} *)
